PROGRAM MAIN
VAR
	_defaultContext : DefaultContext;
	_cylinderBaseTests : CylinderBaseTestContext;
	_doubleCylinderBaseTests : DoubleCylinderBaseTestContext;
		

	_cylinderTests : CylinderTestContext;
	_doubleCylinderTests : DoubleCylinderTestContext;
END_VAR

_defaultContext.Run();
_cylinderTests.ProbeRun();
_doubleCylinderTests.ProbeRun();

_cylinderBaseTests.ProbeRun();
_doublecylinderBaseTests.ProbeRun();

END_PROGRAM

(* stored: Version 1.1.0.1, ProductVersion 3.1.4024.10
   POU MAIN: Id {6d949533-a6b9-47e3-b85f-8c626bcf836e}, SpecialFunc None *)
